Fanuc KAREL source: KA00025.KL

PROGRAM KA00025
%NOLOCKGROUP
VAR
  SRC: BOOLEAN
  DST: INTEGER
BEGIN
  SRC = TRUE
  DST = SRC
END KA00025
